Staubli VAL3: ManyMoves.pjx

--- ManyMoves.pjx ---
Parameters version=s7.5.3 stackSize=5000 millimeterUnit=true
Program file=MoveJoint.pgx
Program file=MoveLine.pgx
Program file=start.pgx
Program file=stop.pgx
Program file=main.pgx
Data file=ManyMoves.dtx

--- ManyMoves.dtx ---
mdesc mNomSpeed
frame fFrame1 = {x=1234.570, y=-98.765, z=50.500, rx=-0.000, ry=0.000, rz=30.000, fatherId=world[0]}
dio Input[16]
  [0] = {link=BasicIO-1\%I0}
  [1] = {link=BasicIO-1\%I1}
  [2] = {link=BasicIO-1\%I2}
  [3] = {link=BasicIO-1\%I3}
  [4] = {link=BasicIO-1\%I4}
  [5] = {link=BasicIO-1\%I5}
  [6] = {link=BasicIO-1\%I6}
  [7] = {link=BasicIO-1\%I7}
  [8] = {link=BasicIO-1\%I8}
  [9] = {link=BasicIO-1\%I9}
  [10] = {link=BasicIO-1\%I10}
  [11] = {link=BasicIO-1\%I11}
  [12] = {link=BasicIO-1\%I12}
  [13] = {link=BasicIO-1\%I13}
  [14] = {link=BasicIO-1\%I14}
  [15] = {link=BasicIO-1\%I15}
dio Output[16]
  [0] = {link=BasicIO-1\%Q0}
  [1] = {link=BasicIO-1\%Q1}
  [2] = {link=BasicIO-1\%Q2}
  [3] = {link=BasicIO-1\%Q3}
  [4] = {link=BasicIO-1\%Q4}
  [5] = {link=BasicIO-1\%Q5}
  [6] = {link=BasicIO-1\%Q6}
  [7] = {link=BasicIO-1\%Q7}
  [8] = {link=BasicIO-1\%Q8}
  [9] = {link=BasicIO-1\%Q9}
  [10] = {link=BasicIO-1\%Q10}
  [11] = {link=BasicIO-1\%Q11}
  [12] = {link=BasicIO-1\%Q12}
  [13] = {link=BasicIO-1\%Q13}
  [14] = {link=BasicIO-1\%Q14}
  [15] = {link=BasicIO-1\%Q15}
tool tCurrentTool = {x=10.000, y=20.000, z=150.000, rx=-0.000, ry=0.000, rz=-0.000, fatherId=flange[0], ioLink=ValveIO/valve1}
mdesc mCurrentSpeed
pointRs pPointRs = {fatherId=fFrame1[0]}
pointRs pPointRs2 = {fatherId=fFrame1[0]}

--- main.pgx ---
program main()
begin
  close(tCurrentTool)
  pPointRs.config.shoulder = lefty
  pPointRs2.config.shoulder = lefty
  mCurrentSpeed.tvel = 100.00
  mCurrentSpeed.blend = joint
  mCurrentSpeed.reach = 0.010
  mCurrentSpeed.leave = 0.010
  // Program ManyMoves start
  // Program generated by RoboDK v6.0.7 for Staubli TP80 on XX/XX/XXXX 18:00:00
  // Using nominal kinematics.
  mCurrentSpeed.tvel = 500.000
  call MoveJoint(10.00000,-20.00000,50.00000,30.00000)
  call MoveLine(-638.084,504.480,372.034,136.262,30.757,-130.375)
  call MoveJoint(30.00000,25.00000,80.00000,-45.00000)
  // Linear movement using joint targets is not supported. Change the target type to cartesian or use a joint movement.
  call MoveJoint(10.00000,-20.00000,50.00000,30.00000)
  call MoveLine(-628.084,494.480,374.034,136.262,30.757,-130.375)
  call MoveJoint(30.00000,25.00000,80.00000,-45.00000)
  // Linear movement using joint targets is not supported. Change the target type to cartesian or use a joint movement.
  call MoveJoint(10.00000,-20.00000,50.00000,30.00000)
  call MoveLine(-618.084,484.480,376.034,136.262,30.757,-130.375)
  call MoveJoint(30.00000,25.00000,80.00000,-45.00000)
  // Linear movement using joint targets is not supported. Change the target type to cartesian or use a joint movement.
  call MoveJoint(10.00000,-20.00000,50.00000,30.00000)
  call MoveLine(-608.084,474.480,378.034,136.262,30.757,-130.375)
  call MoveJoint(30.00000,25.00000,80.00000,-45.00000)
  // Linear movement using joint targets is not supported. Change the target type to cartesian or use a joint movement.
  call MoveJoint(10.00000,-20.00000,50.00000,30.00000)
  call MoveLine(-598.084,464.480,380.034,136.262,30.757,-130.375)
  call MoveJoint(30.00000,25.00000,80.00000,-45.00000)
  // Linear movement using joint targets is not supported. Change the target type to cartesian or use a joint movement.
  call MoveJoint(10.00000,-20.00000,50.00000,30.00000)
  call MoveLine(-588.084,454.480,382.034,136.262,30.757,-130.375)
  call MoveJoint(30.00000,25.00000,80.00000,-45.00000)
  // Linear movement using joint targets is not supported. Change the target type to cartesian or use a joint movement.
  call MoveJoint(10.00000,-20.00000,50.00000,30.00000)
  call MoveLine(-578.084,444.480,384.034,136.262,30.757,-130.375)
  call MoveJoint(30.00000,25.00000,80.00000,-45.00000)
  // Linear movement using joint targets is not supported. Change the target type to cartesian or use a joint movement.
  call MoveJoint(10.00000,-20.00000,50.00000,30.00000)
  call MoveLine(-568.084,434.480,386.034,136.262,30.757,-130.375)
  call MoveJoint(30.00000,25.00000,80.00000,-45.00000)
  // Linear movement using joint targets is not supported. Change the target type to cartesian or use a joint movement.
  call MoveJoint(10.00000,-20.00000,50.00000,30.00000)
  call MoveLine(-558.084,424.480,388.034,136.262,30.757,-130.375)
  call MoveJoint(30.00000,25.00000,80.00000,-45.00000)
  // Linear movement using joint targets is not supported. Change the target type to cartesian or use a joint movement.
  call MoveJoint(10.00000,-20.00000,50.00000,30.00000)
  call MoveLine(-548.084,414.480,390.034,136.262,30.757,-130.375)
  call MoveJoint(30.00000,25.00000,80.00000,-45.00000)
  // Linear movement using joint targets is not supported. Change the target type to cartesian or use a joint movement.

  waitEndMove()
  // Program ManyMoves end

end

--- start.pgx ---
program start()
begin
  call main()
end

--- MoveJoint.pgx ---
program MoveJoint(num x_nJ1, num x_nJ2, num x_nJ3, num x_nJ4)
  local joint l_jJoint
begin
  l_jJoint.j1 = x_nJ1
  l_jJoint.j2 = x_nJ2
  l_jJoint.j3 = x_nJ3
  l_jJoint.j4 = x_nJ4
  movej(l_jJoint,tCurrentTool ,mCurrentSpeed)
end

--- MoveLine.pgx ---
program MoveLine(num x_nX, num x_nY, num x_nZ, num x_nRx, num x_nRy, num x_nRz)
begin
  pPointRs.trsf.x = x_nX
  pPointRs.trsf.y = x_nY
  pPointRs.trsf.z = x_nZ
  pPointRs.trsf.rx = x_nRx
  pPointRs.trsf.ry = x_nRy
  pPointRs.trsf.rz = x_nRz
  movel(pPointRs,tCurrentTool,mCurrentSpeed)
end

--- stop.pgx ---
program stop()
begin
end
